Fanuc KAREL source: kt00129.KL

-- PROVISIONAL review KL for V1013-1; original PC SHA256 e1232820cf35ac1bf899cb7b82ff67e1b4625c57b88a8f263073c8e44dc0464a
-- Incomplete behavior may be omitted. Consult companion uncertainty JSON. Do not deploy.
PROGRAM KT00129
%NOLOCKGROUP
VAR
  I1 : INTEGER
  I2 : INTEGER
  OUT : INTEGER
BEGIN
  -- UNRESOLVED_PC offsets 5-16; opcodes 2E,23
  -- UNRESOLVED_PC offsets 21-32; opcodes 2E,23
  -- UNRESOLVED_PC offsets 37-48; opcodes 2E,23
  -- UNRESOLVED_PC offsets 53-64; opcodes 2E,23
  -- UNRESOLVED_PC offsets 69-88; opcodes 21,21,55,23
  -- UNRESOLVED_PC offsets 93-97; opcodes 7F
END KT00129
